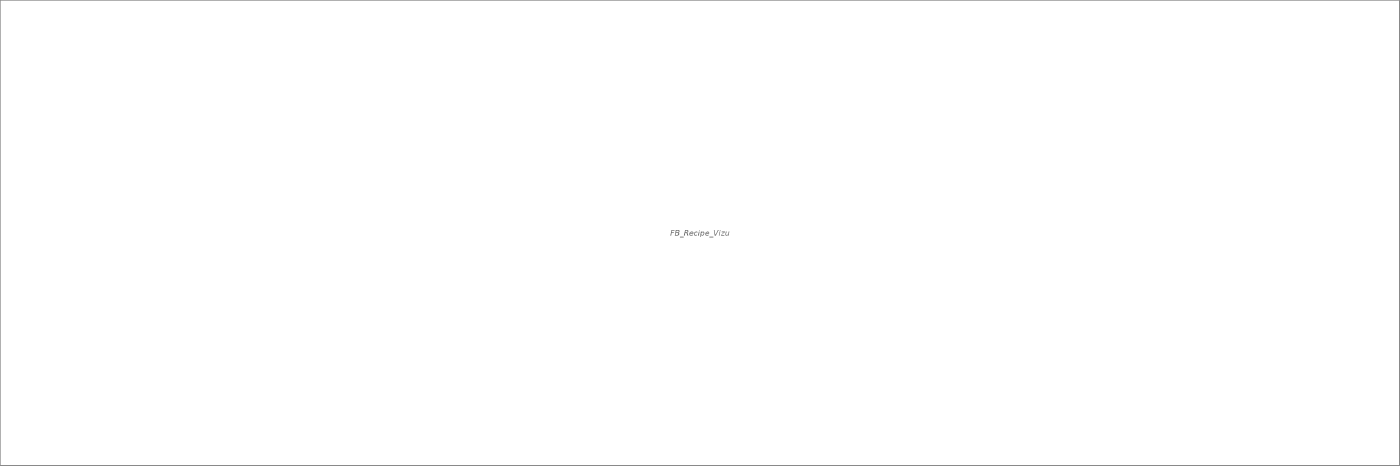
VISUALIZATION Vis_Recipe_Tab  // 1850x617
    TabControl (0,0 1850x617), frame switch variable: prg_Call_Recipe_Slow.iRecipeSwitchFrameVar
        shows FB_Recipe_Vizu(fb_Recipe := GVL_Recipe.fbRecipe[E_Recipe_Name.R_All])
        shows FB_Recipe_Vizu(fb_Recipe := GVL_Recipe.fbRecipe[E_Recipe_Name.R_Device_Dough1])
        shows FB_Recipe_Vizu(fb_Recipe := GVL_Recipe.fbRecipe[E_Recipe_Name.R_Device_Dough2])
        shows FB_Recipe_Vizu(fb_Recipe := GVL_Recipe.fbRecipe[E_Recipe_Name.R_Device_Dough3])
        shows FB_Recipe_Vizu(fb_Recipe := GVL_Recipe.fbRecipe[E_Recipe_Name.R_Device_Dough4])
        shows FB_Recipe_Vizu(fb_Recipe := GVL_Recipe.fbRecipe[E_Recipe_Name.R_CheesyBites])
        shows FB_Recipe_Vizu(fb_Recipe := GVL_Recipe.fbRecipe[E_Recipe_Name.R_CheesyCut])
        shows FB_Recipe_Vizu(fb_Recipe := GVL_Recipe.fbRecipe[E_Recipe_Name.R_Cream])
        shows FB_Recipe_Vizu(fb_Recipe := GVL_Recipe.fbRecipe[E_Recipe_Name.R_Crown])
        shows FB_Recipe_Vizu(fb_Recipe := GVL_Recipe.fbRecipe[E_Recipe_Name.R_Flour])
        shows FB_Recipe_Vizu(fb_Recipe := GVL_Recipe.fbRecipe[E_Recipe_Name.R_Mozzarella])
        shows FB_Recipe_Vizu(fb_Recipe := GVL_Recipe.fbRecipe[E_Recipe_Name.R_Open1])
        shows FB_Recipe_Vizu(fb_Recipe := GVL_Recipe.fbRecipe[E_Recipe_Name.R_Open2])
        shows FB_Recipe_Vizu(fb_Recipe := GVL_Recipe.fbRecipe[E_Recipe_Name.R_Open3])
        shows FB_Recipe_Vizu(fb_Recipe := GVL_Recipe.fbRecipe[E_Recipe_Name.R_Open4])
        shows FB_Recipe_Vizu(fb_Recipe := GVL_Recipe.fbRecipe[E_Recipe_Name.R_Wet])
        shows FB_Recipe_Vizu(fb_Recipe := GVL_Recipe.fbRecipe[E_Recipe_Name.R_Wrap])
        shows FB_Recipe_Vizu(fb_Recipe := GVL_Recipe.fbRecipe[E_Recipe_Name.R_Sesame])
        shows FB_Recipe_Vizu(fb_Recipe := GVL_Recipe.fbRecipe[E_Recipe_Name.R_Piston_Settings])
        [0]: TabTitle=All
        [1]: TabTitle=Device 1
        [2]: TabTitle=Device 2
        [3]: TabTitle=Device 3
        [4]: TabTitle=Device 4
        [5]: TabTitle=Cheesy Bites
        [6]: TabTitle=Cheesy Cut
        [7]: TabTitle=Cream
        [8]: TabTitle=Crown
        [9]: TabTitle=Flour
        [10]: TabTitle=Mozza
        [11]: TabTitle=Open1
        [12]: TabTitle=Open2
        [13]: TabTitle=Open3
        [14]: TabTitle=Open4
        [15]: TabTitle=Wet
        [16]: TabTitle=Wrap
        [17]: TabTitle=Sesame
        [18]: TabTitle=Piston Param
END_VISUALIZATION

(* stored: Version 1.1.0.1, ProductVersion 3.1.4024.12
   Visu Vis_Recipe_Tab: Id {d84762c1-01a5-46ba-8e85-524383057f09} *)
